Universal Robots URScript: horizontal_swab_path 4.script

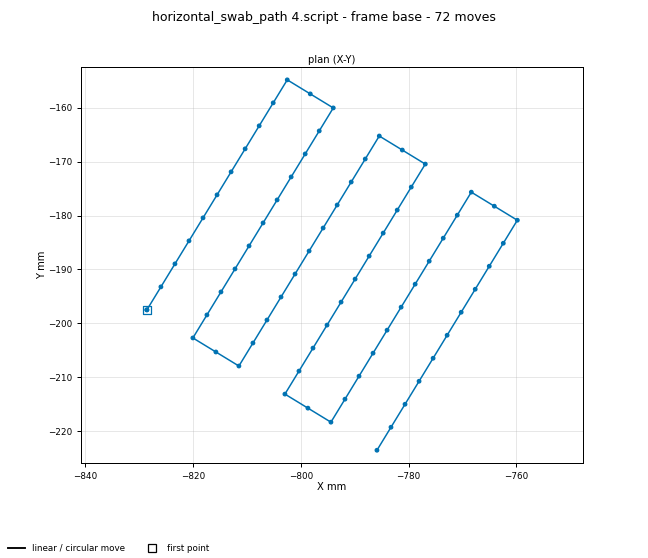
[picture p0: tool path of horizontal_swab_path 4.script in frame base, 72 of 72 moves have a stored position in this frame; points joined in program order, loops and branches not executed]
def horizontal_swab_path():

  # Move to first swab point perpendicular
  movel(p[-0.82856417, -0.19749532, 0.03086437, -0.84988534, -3.02427359, 0.03157596], a=0.2000, v=0.0300, r=0.0000)

  # Incline tool while keeping TCP XYZ fixed
  movel(p[-0.82856417, -0.19749532, 0.03086437, -0.65161072, -2.28357471, -0.24197279], a=0.1000, v=0.0150, r=0.0000)
  # Horizontal waypoint 1
  movel(p[-0.82595991, -0.19322818, 0.03076760, -0.65161072, -2.28357471, -0.24197279], a=0.1500, v=0.0200, r=0.0000)
  # Horizontal waypoint 2
  movel(p[-0.82335565, -0.18896104, 0.03067083, -0.65161072, -2.28357471, -0.24197279], a=0.1500, v=0.0200, r=0.0000)
  # Horizontal waypoint 3
  movel(p[-0.82075138, -0.18469391, 0.03057406, -0.65161072, -2.28357471, -0.24197279], a=0.1500, v=0.0200, r=0.0000)
  # Horizontal waypoint 4
  movel(p[-0.81814712, -0.18042677, 0.03047728, -0.65161072, -2.28357471, -0.24197279], a=0.1500, v=0.0200, r=0.0000)
  # Horizontal waypoint 5
  movel(p[-0.81554286, -0.17615963, 0.03038051, -0.65161072, -2.28357471, -0.24197279], a=0.1500, v=0.0200, r=0.0000)
  # Horizontal waypoint 6
  movel(p[-0.81293860, -0.17189250, 0.03028374, -0.65161072, -2.28357471, -0.24197279], a=0.1500, v=0.0200, r=0.0000)
  # Horizontal waypoint 7
  movel(p[-0.81033434, -0.16762536, 0.03018697, -0.65161072, -2.28357471, -0.24197279], a=0.1500, v=0.0200, r=0.0000)
  # Horizontal waypoint 8
  movel(p[-0.80773007, -0.16335822, 0.03009020, -0.65161072, -2.28357471, -0.24197279], a=0.1500, v=0.0200, r=0.0000)
  # Horizontal waypoint 9
  movel(p[-0.80512581, -0.15909109, 0.02999342, -0.65161072, -2.28357471, -0.24197279], a=0.1500, v=0.0200, r=0.0000)
  # Horizontal waypoint 10
  movel(p[-0.80252155, -0.15482395, 0.02989665, -0.65161072, -2.28357471, -0.24197279], a=0.1500, v=0.0200, r=0.0000)
  # Horizontal waypoint 11
  movel(p[-0.79825340, -0.15742822, 0.02992379, -0.65161072, -2.28357471, -0.24197279], a=0.1500, v=0.0200, r=0.0000)
  # Horizontal waypoint 12
  movel(p[-0.79398526, -0.16003248, 0.02995092, -0.65161072, -2.28357471, -0.24197279], a=0.1500, v=0.0200, r=0.0000)
  # Horizontal waypoint 13
  movel(p[-0.79658952, -0.16429962, 0.03004769, -0.65161072, -2.28357471, -0.24197279], a=0.1500, v=0.0200, r=0.0000)
  # Horizontal waypoint 14
  movel(p[-0.79919378, -0.16856675, 0.03014446, -0.65161072, -2.28357471, -0.24197279], a=0.1500, v=0.0200, r=0.0000)
  # Horizontal waypoint 15
  movel(p[-0.80179804, -0.17283389, 0.03024124, -0.65161072, -2.28357471, -0.24197279], a=0.1500, v=0.0200, r=0.0000)
  # Horizontal waypoint 16
  movel(p[-0.80440230, -0.17710102, 0.03033801, -0.65161072, -2.28357471, -0.24197279], a=0.1500, v=0.0200, r=0.0000)
  # Horizontal waypoint 17
  movel(p[-0.80700657, -0.18136816, 0.03043478, -0.65161072, -2.28357471, -0.24197279], a=0.1500, v=0.0200, r=0.0000)
  # Horizontal waypoint 18
  movel(p[-0.80961083, -0.18563530, 0.03053155, -0.65161072, -2.28357471, -0.24197279], a=0.1500, v=0.0200, r=0.0000)
  # Horizontal waypoint 19
  movel(p[-0.81221509, -0.18990243, 0.03062833, -0.65161072, -2.28357471, -0.24197279], a=0.1500, v=0.0200, r=0.0000)
  # Horizontal waypoint 20
  movel(p[-0.81481935, -0.19416957, 0.03072510, -0.65161072, -2.28357471, -0.24197279], a=0.1500, v=0.0200, r=0.0000)
  # Horizontal waypoint 21
  movel(p[-0.81742362, -0.19843671, 0.03082187, -0.65161072, -2.28357471, -0.24197279], a=0.1500, v=0.0200, r=0.0000)
  # Horizontal waypoint 22
  movel(p[-0.82002788, -0.20270384, 0.03091864, -0.65161072, -2.28357471, -0.24197279], a=0.1500, v=0.0200, r=0.0000)
  # Horizontal waypoint 23
  movel(p[-0.81575973, -0.20530811, 0.03094578, -0.65161072, -2.28357471, -0.24197279], a=0.1500, v=0.0200, r=0.0000)
  # Horizontal waypoint 24
  movel(p[-0.81149158, -0.20791237, 0.03097291, -0.65161072, -2.28357471, -0.24197279], a=0.1500, v=0.0200, r=0.0000)
  # Horizontal waypoint 25
  movel(p[-0.80888732, -0.20364523, 0.03087614, -0.65161072, -2.28357471, -0.24197279], a=0.1500, v=0.0200, r=0.0000)
  # Horizontal waypoint 26
  movel(p[-0.80628306, -0.19937810, 0.03077937, -0.65161072, -2.28357471, -0.24197279], a=0.1500, v=0.0200, r=0.0000)
  # Horizontal waypoint 27
  movel(p[-0.80367880, -0.19511096, 0.03068260, -0.65161072, -2.28357471, -0.24197279], a=0.1500, v=0.0200, r=0.0000)
  # Horizontal waypoint 28
  movel(p[-0.80107454, -0.19084382, 0.03058582, -0.65161072, -2.28357471, -0.24197279], a=0.1500, v=0.0200, r=0.0000)
  # Horizontal waypoint 29
  movel(p[-0.79847027, -0.18657669, 0.03048905, -0.65161072, -2.28357471, -0.24197279], a=0.1500, v=0.0200, r=0.0000)
  # Horizontal waypoint 30
  movel(p[-0.79586601, -0.18230955, 0.03039228, -0.65161072, -2.28357471, -0.24197279], a=0.1500, v=0.0200, r=0.0000)
  # Horizontal waypoint 31
  movel(p[-0.79326175, -0.17804242, 0.03029551, -0.65161072, -2.28357471, -0.24197279], a=0.1500, v=0.0200, r=0.0000)
  # Horizontal waypoint 32
  movel(p[-0.79065749, -0.17377528, 0.03019873, -0.65161072, -2.28357471, -0.24197279], a=0.1500, v=0.0200, r=0.0000)
  # Horizontal waypoint 33
  movel(p[-0.78805322, -0.16950814, 0.03010196, -0.65161072, -2.28357471, -0.24197279], a=0.1500, v=0.0200, r=0.0000)
  # Horizontal waypoint 34
  movel(p[-0.78544896, -0.16524100, 0.03000519, -0.65161072, -2.28357471, -0.24197279], a=0.1500, v=0.0200, r=0.0000)
  # Horizontal waypoint 35
  movel(p[-0.78118082, -0.16784527, 0.03003232, -0.65161072, -2.28357471, -0.24197279], a=0.1500, v=0.0200, r=0.0000)
  # Horizontal waypoint 36
  movel(p[-0.77691267, -0.17044953, 0.03005946, -0.65161072, -2.28357471, -0.24197279], a=0.1500, v=0.0200, r=0.0000)
  # Horizontal waypoint 37
  movel(p[-0.77951693, -0.17471667, 0.03015623, -0.65161072, -2.28357471, -0.24197279], a=0.1500, v=0.0200, r=0.0000)
  # Horizontal waypoint 38
  movel(p[-0.78212119, -0.17898380, 0.03025300, -0.65161072, -2.28357471, -0.24197279], a=0.1500, v=0.0200, r=0.0000)
  # Horizontal waypoint 39
  movel(p[-0.78472546, -0.18325094, 0.03034978, -0.65161072, -2.28357471, -0.24197279], a=0.1500, v=0.0200, r=0.0000)
  # Horizontal waypoint 40
  movel(p[-0.78732972, -0.18751808, 0.03044655, -0.65161072, -2.28357471, -0.24197279], a=0.1500, v=0.0200, r=0.0000)
  # Horizontal waypoint 41
  movel(p[-0.78993398, -0.19178521, 0.03054332, -0.65161072, -2.28357471, -0.24197279], a=0.1500, v=0.0200, r=0.0000)
  # Horizontal waypoint 42
  movel(p[-0.79253824, -0.19605235, 0.03064009, -0.65161072, -2.28357471, -0.24197279], a=0.1500, v=0.0200, r=0.0000)
  # Horizontal waypoint 43
  movel(p[-0.79514251, -0.20031949, 0.03073687, -0.65161072, -2.28357471, -0.24197279], a=0.1500, v=0.0200, r=0.0000)
  # Horizontal waypoint 44
  movel(p[-0.79774677, -0.20458662, 0.03083364, -0.65161072, -2.28357471, -0.24197279], a=0.1500, v=0.0200, r=0.0000)
  # Horizontal waypoint 45
  movel(p[-0.80035103, -0.20885376, 0.03093041, -0.65161072, -2.28357471, -0.24197279], a=0.1500, v=0.0200, r=0.0000)
  # Horizontal waypoint 46
  movel(p[-0.80295529, -0.21312090, 0.03102718, -0.65161072, -2.28357471, -0.24197279], a=0.1500, v=0.0200, r=0.0000)
  # Horizontal waypoint 47
  movel(p[-0.79868715, -0.21572516, 0.03105432, -0.65161072, -2.28357471, -0.24197279], a=0.1500, v=0.0200, r=0.0000)
  # Horizontal waypoint 48
  movel(p[-0.79441900, -0.21832942, 0.03108145, -0.65161072, -2.28357471, -0.24197279], a=0.1500, v=0.0200, r=0.0000)
  # Horizontal waypoint 49
  movel(p[-0.79181474, -0.21406229, 0.03098468, -0.65161072, -2.28357471, -0.24197279], a=0.1500, v=0.0200, r=0.0000)
  # Horizontal waypoint 50
  movel(p[-0.78921047, -0.20979515, 0.03088791, -0.65161072, -2.28357471, -0.24197279], a=0.1500, v=0.0200, r=0.0000)
  # Horizontal waypoint 51
  movel(p[-0.78660621, -0.20552801, 0.03079114, -0.65161072, -2.28357471, -0.24197279], a=0.1500, v=0.0200, r=0.0000)
  # Horizontal waypoint 52
  movel(p[-0.78400195, -0.20126088, 0.03069436, -0.65161072, -2.28357471, -0.24197279], a=0.1500, v=0.0200, r=0.0000)
  # Horizontal waypoint 53
  movel(p[-0.78139769, -0.19699374, 0.03059759, -0.65161072, -2.28357471, -0.24197279], a=0.1500, v=0.0200, r=0.0000)
  # Horizontal waypoint 54
  movel(p[-0.77879343, -0.19272660, 0.03050082, -0.65161072, -2.28357471, -0.24197279], a=0.1500, v=0.0200, r=0.0000)
  # Horizontal waypoint 55
  movel(p[-0.77618916, -0.18845947, 0.03040405, -0.65161072, -2.28357471, -0.24197279], a=0.1500, v=0.0200, r=0.0000)
  # Horizontal waypoint 56
  movel(p[-0.77358490, -0.18419233, 0.03030727, -0.65161072, -2.28357471, -0.24197279], a=0.1500, v=0.0200, r=0.0000)
  # Horizontal waypoint 57
  movel(p[-0.77098064, -0.17992520, 0.03021050, -0.65161072, -2.28357471, -0.24197279], a=0.1500, v=0.0200, r=0.0000)
  # Horizontal waypoint 58
  movel(p[-0.76837638, -0.17565806, 0.03011373, -0.65161072, -2.28357471, -0.24197279], a=0.1500, v=0.0200, r=0.0000)
  # Horizontal waypoint 59
  movel(p[-0.76410823, -0.17826232, 0.03014086, -0.65161072, -2.28357471, -0.24197279], a=0.1500, v=0.0200, r=0.0000)
  # Horizontal waypoint 60
  movel(p[-0.75984008, -0.18086659, 0.03016800, -0.65161072, -2.28357471, -0.24197279], a=0.1500, v=0.0200, r=0.0000)
  # Horizontal waypoint 61
  movel(p[-0.76244435, -0.18513372, 0.03026477, -0.65161072, -2.28357471, -0.24197279], a=0.1500, v=0.0200, r=0.0000)
  # Horizontal waypoint 62
  movel(p[-0.76504861, -0.18940086, 0.03036154, -0.65161072, -2.28357471, -0.24197279], a=0.1500, v=0.0200, r=0.0000)
  # Horizontal waypoint 63
  movel(p[-0.76765287, -0.19366800, 0.03045831, -0.65161072, -2.28357471, -0.24197279], a=0.1500, v=0.0200, r=0.0000)
  # Horizontal waypoint 64
  movel(p[-0.77025713, -0.19793513, 0.03055509, -0.65161072, -2.28357471, -0.24197279], a=0.1500, v=0.0200, r=0.0000)
  # Horizontal waypoint 65
  movel(p[-0.77286139, -0.20220227, 0.03065186, -0.65161072, -2.28357471, -0.24197279], a=0.1500, v=0.0200, r=0.0000)
  # Horizontal waypoint 66
  movel(p[-0.77546566, -0.20646940, 0.03074863, -0.65161072, -2.28357471, -0.24197279], a=0.1500, v=0.0200, r=0.0000)
  # Horizontal waypoint 67
  movel(p[-0.77806992, -0.21073654, 0.03084540, -0.65161072, -2.28357471, -0.24197279], a=0.1500, v=0.0200, r=0.0000)
  # Horizontal waypoint 68
  movel(p[-0.78067418, -0.21500368, 0.03094218, -0.65161072, -2.28357471, -0.24197279], a=0.1500, v=0.0200, r=0.0000)
  # Horizontal waypoint 69
  movel(p[-0.78327844, -0.21927081, 0.03103895, -0.65161072, -2.28357471, -0.24197279], a=0.1500, v=0.0200, r=0.0000)
  # Horizontal waypoint 70
  movel(p[-0.78588271, -0.22353795, 0.03113572, -0.65161072, -2.28357471, -0.24197279], a=0.1500, v=0.0200, r=0.0000)

end
